// TIA Portal V21 export
DATA_BLOCK "IDB_LadOpenBranch"   // DB21
// stored: InstanceOfName FB_LadOpenBranch, InstanceOfType FB
"FB_LadOpenBranch"
   // VAR_INPUT
   //    Start : Bool;
   //    Stop : Bool;
   // END_VAR
   // VAR_OUTPUT
   //    CoilA : Bool;
   //    CoilB : Bool;
   //    CoilC : Bool;
   //    BranchOut : Bool;
   //    StopLatched : Bool;
   // END_VAR
   // VAR
   //    StartCount : Int;
   // END_VAR
BEGIN
END_DATA_BLOCK
